PROGRAM main
  VAR
    step0 : BOOL;
    step1 : BOOL;
    step2 : BOOL;
    step3 : BOOL;
    step4 : BOOL;
    T1 : BOOL;
    T2 : BOOL;
    T3 : BOOL;
    led_rosso : BOOL;
    led_giallo : BOOL;
    led_verde : BOOL;
    start : BOOL;
    TON0 : TON;
    TON1 : TON;
    TON2 : TON;
  END_VAR
  VAR_INPUT
  END_VAR

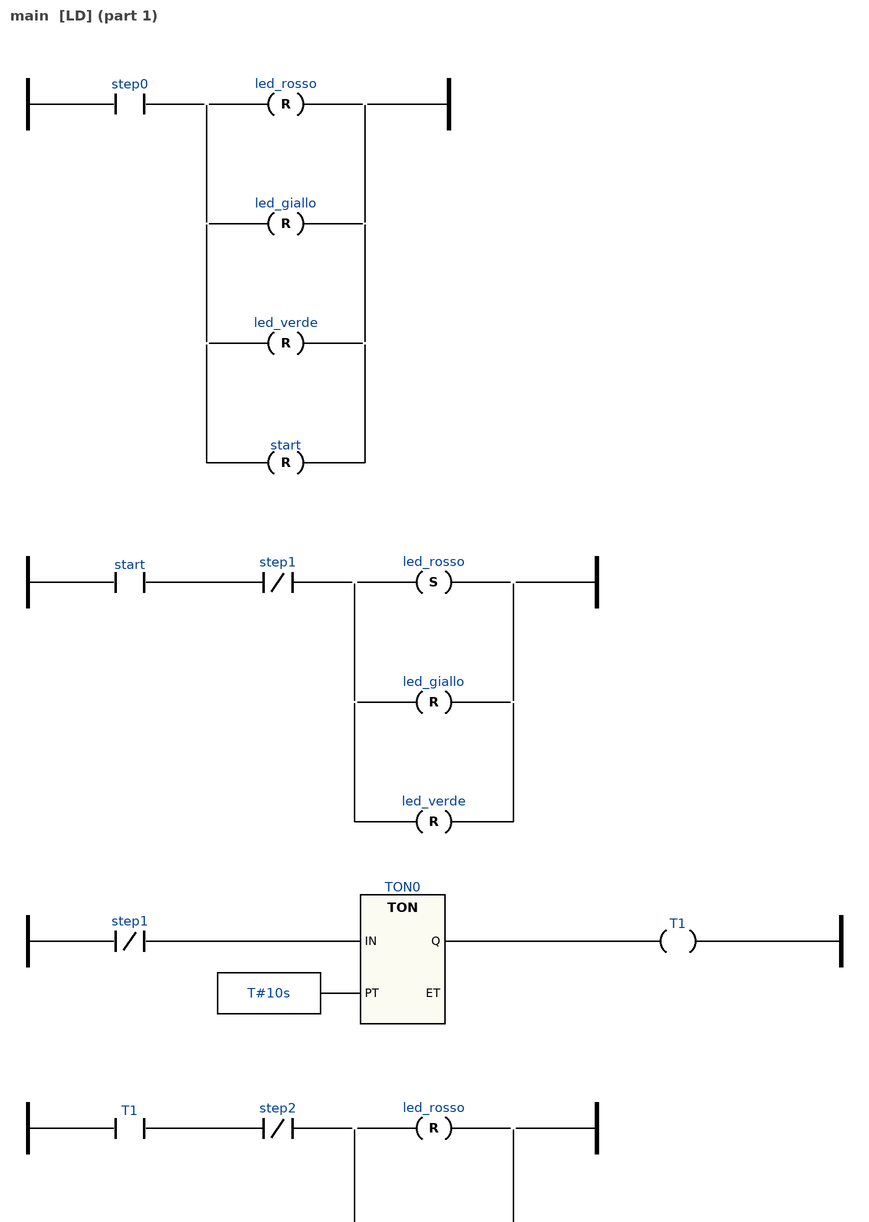
(* LD diagram, written out as Structured Text *)
IF step0 THEN led_rosso := FALSE; END_IF;
IF step0 THEN led_giallo := FALSE; END_IF;
IF step0 THEN led_verde := FALSE; END_IF;
IF step0 THEN start := FALSE; END_IF;
IF start AND NOT step1 THEN led_rosso := TRUE; END_IF;
IF start AND NOT step1 THEN led_giallo := FALSE; END_IF;
IF start AND NOT step1 THEN led_verde := FALSE; END_IF;
TON0(IN := NOT step1, PT := T#10s);
T1 := TON0.Q;
IF T1 AND NOT step2 THEN led_rosso := FALSE; END_IF;
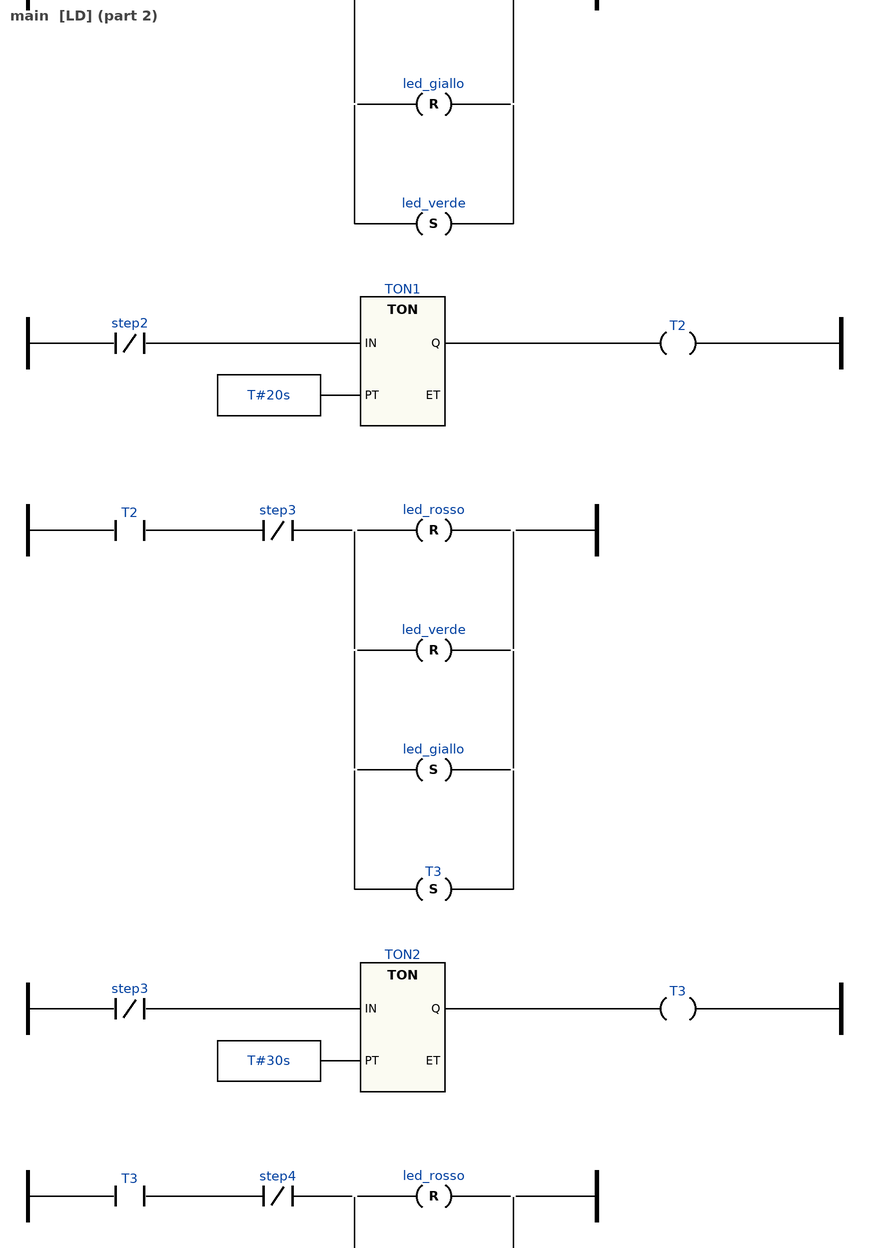
IF T1 AND NOT step2 THEN led_giallo := FALSE; END_IF;
IF T1 AND NOT step2 THEN led_verde := TRUE; END_IF;
TON1(IN := NOT step2, PT := T#20s);
T2 := TON1.Q;
IF T2 AND NOT step3 THEN led_rosso := FALSE; END_IF;
IF T2 AND NOT step3 THEN led_verde := FALSE; END_IF;
IF T2 AND NOT step3 THEN led_giallo := TRUE; END_IF;
IF T2 AND NOT step3 THEN T3 := TRUE; END_IF;
TON2(IN := NOT step3, PT := T#30s);
T3 := TON2.Q;
IF T3 AND NOT step4 THEN led_rosso := FALSE; END_IF;
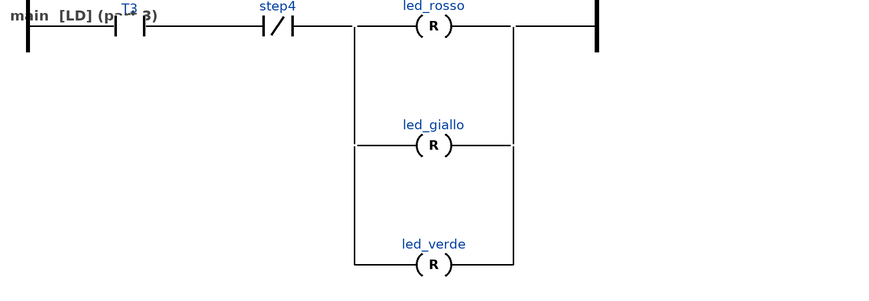
IF T3 AND NOT step4 THEN led_giallo := FALSE; END_IF;
IF T3 AND NOT step4 THEN led_verde := FALSE; END_IF;
END_PROGRAM
